PROGRAM MAIN
VAR
	fbMotionSystem	: FB_MotionSystem;
	nState			: UDINT;
END_VAR

// Main program: start up the system, enable it, then run the exercise.
CASE nState OF
	0:	nState := 1;
	1:	IF fbMotionSystem.Startup() THEN
			nState := 30;
		END_IF
	30:	IF fbMotionSystem.Starting(bReset := FALSE) THEN
			nState := 40;
		END_IF
	40:	fbMotionSystem.Execute();	// movers drive between the stations
END_CASE

fbMotionSystem.Cycle();

END_PROGRAM

(* stored: Version 1.1.0.1
   POU MAIN: Id {2767b9cb-02c7-4e83-9bc7-d611a48e2aad} *)
